// TIA Portal project "000_empty" (V21)

(* hardware
DEVICE "PLC_1"  S7-1500 station
   slot 0: "Rail_0"  Rack  6ES7 590-1***0-0AA0
   slot 1: "PLC_1"  CPU 1513-1 PN  6ES7 513-1AL02-0AB0  V2.9
      slot 3: "CPU display_1"  6ES7591-1AA00-0AA0
      slot 32768: "PROFINET interface_1"  X1
         slot 32769: "Port_1"  X1 P1
         slot 32770: "Port_2"  X1 P2
      slot 34817: "Virtual CP interface port_1"  Virtual CP interface port  Virtual CP interface port
*)

// ===== PLC "PLC_1"  CPU 1513-1 PN =====

VAR_GLOBAL   // PLC tag table "Default tag table"
   "tBool" AT %M0.0 : Bool;
   "tBool2" AT %M0.1 : Bool;
   "tInt" AT %MW2 : Int;
   "tDInt" AT %MD4 : DInt;
   "tReal" AT %MD8 : Real;
   "tWord" AT %MW12 : Word;
   "tByte" AT %MB14 : Byte;
   "tDWord" AT %MD16 : DWord;
   "tTime" AT %MD20 : Time;
   "tIn" AT %I0.0 : Bool;
   "tOut" AT %Q0.0 : Bool;
   "tUInt" AT %MW24 : UInt;
   "tLReal" AT %MD26 : LReal;
   "Tag_1" AT %MW100 : Word;
   "Tag_2" AT %M10.3 : Bool;
   "Tag_3" AT %Q1.0 : Bool;
   "Tag_4" AT %I1.0 : Bool;
   "Tag_5" AT %MD104 : DWord;
   "Tag_6" AT %MB110 : Byte;
   "Tag_7" AT %IW0 : Word;
   "Tag_8" AT %QW0 : Word;
END_VAR

VAR_GLOBAL CONSTANT   // PLC tag table "Default tag table"
   "MAX_COUNT" : Int := 100;
   "GAIN" : Real := 2.5;
   "TXT" : String := 'abc';
END_VAR

TYPE "UDT_Motor"
   STRUCT
      Running : Bool;   // Motor on
      Speed : Real := 1500.0;   // Speed setpoint
      Count : Int := 7;
   END_STRUCT;
END_TYPE

DATA_BLOCK "DB_Global"   // DB1
{ S7_Optimized_Access := 'TRUE' }
   VAR
      xBool : Bool := TRUE;   // Bool comment
      iInt : Int := 42;
      rReal : Real := 3.5;   // Real comment
      aInt : Array[0..3] of Int;
      sData : Struct
         "a" : Bool;
         "b" : DInt := -5;
      END_STRUCT;
   END_VAR
BEGIN
   aInt[1] := 11;
END_DATA_BLOCK

DATA_BLOCK "FB_Empty_DB"   // DB2
{ S7_Optimized_Access := 'TRUE' }
VERSION : 0.1
// stored: InstanceOfName FB_Empty
"FB_Empty"
BEGIN
END_DATA_BLOCK

DATA_BLOCK "DB_Motor"   // DB4
{ S7_Optimized_Access := 'TRUE' }
   VAR
      motor : "UDT_Motor";
   END_VAR
BEGIN
   motor.Speed := 750.0;
END_DATA_BLOCK

DATA_BLOCK "FB_Iface_DB"   // DB5
{ S7_Optimized_Access := 'TRUE' }
VERSION : 0.1
// stored: InstanceOfName FB_Iface
"FB_Iface"
BEGIN
   stInt := 99;
   stBool := TRUE;
END_DATA_BLOCK

DATA_BLOCK "DB_Std"   // DB6
{ S7_Optimized_Access := 'FALSE' }
   VAR
      x : Bool;
      i : Int;
      d : DInt;
      r : Real;
      "by" : Byte;
   END_VAR
BEGIN
END_DATA_BLOCK

DATA_BLOCK "DB_Arr"   // DB7
{ S7_Optimized_Access := 'FALSE' }
   VAR
      "a" : Array[0..9] of Int;
      "b" : Array[0..9] of Int;
      w : Array[0..3] of Word;
      r : Array[0..3] of Real;
      "by" : Array[0..7] of Byte;
      bits : Array[0..15] of Bool;
   END_VAR
BEGIN
END_DATA_BLOCK

// folder: BlockGroup_1

DATA_BLOCK "DB_InGroup"   // DB3
{ S7_Optimized_Access := 'TRUE' }
   VAR
      wWord : Word := 16#00FF;
   END_VAR
BEGIN
END_DATA_BLOCK

// folder: (top level)

FUNCTION_BLOCK "FB_Empty"   // FB1, SCL
{ S7_Optimized_Access := 'TRUE' }
VERSION : 0.1
BEGIN
END_FUNCTION_BLOCK

FUNCTION_BLOCK "FB_Iface"   // FB2, SCL
{ S7_Optimized_Access := 'TRUE' }
VERSION : 0.1
   VAR_INPUT
      iBool : Bool;   // Input bool
      iInt : Int;   // Input int
      iReal : Real;   // Input real
      iArr : Array[0..3] of Int;   // Input array
      iMotor : "UDT_Motor";   // Input UDT
   END_VAR
   VAR_OUTPUT
      oBool : Bool;   // Output bool
      oInt : Int;   // Output int
   END_VAR
   VAR_IN_OUT
      ioReal : Real;   // InOut real
   END_VAR
   VAR
      stInt : Int := 42;   // Static int
      stBool : Bool;   // Static bool comment
   END_VAR
   VAR_TEMP
      tInt : Int;   // Temp int
   END_VAR
   VAR CONSTANT
      cInt : Int := 7;   // Constant int
   END_VAR
BEGIN
   #tInt := #iInt + #cInt;
           #oInt := #tInt;
           #oBool := #iBool;
           #ioReal := #ioReal + #iReal;
END_FUNCTION_BLOCK

FUNCTION_BLOCK "FB_SclCalls"   // FB3, SCL
{ S7_Optimized_Access := 'TRUE' }
VERSION : 0.1
   VAR_INPUT
      start : Bool;
      pt : Time;
   END_VAR
   VAR_OUTPUT
      q : Bool;
      cnt : Int;
   END_VAR
   VAR
      tonInst : TON_TIME;
      tofInst : TOF_TIME;
      tpInst : TP_TIME;
      ctuInst : CTU_INT;
      trig : R_TRIG;
      ftrig : F_TRIG;
      "counter" : Int;
      ifc : "FB_Iface";
   END_VAR
   VAR_TEMP
      r : Real;
      "b" : Bool;
      res : Int;
      tot : Int;
   END_VAR
BEGIN
   #tonInst(IN := #start, PT := #pt);
   #q := #tonInst.Q;
   #tofInst(IN := #start, PT := T#2s);
   #tpInst(IN := #start, PT := #pt, Q => #b);
   #ctuInst(CU := #start, R := FALSE, PV := 10);
   #cnt := #ctuInst.CV;
   #trig(CLK := #start);
   IF #trig.Q THEN
       #counter := 0;
   END_IF;
   #ftrig(CLK := #start);
   #b := #ftrig.Q;
   #ifc(iBool := TRUE, iInt := 2, iReal := 1.0, ioReal := #r);
   #cnt := #ifc.oInt;
   "FB_Iface_DB"(iBool := #start, iInt := #cnt, iReal := #r, ioReal := #r, oInt => #cnt);
   "FC_SclOps"();
   #res := "FC_SclCtl"(n := 5, flag := TRUE, total => #tot);
   #res := "FC_SclCtl"(n := #res, flag := #b, total => #tot);
END_FUNCTION_BLOCK

FUNCTION_BLOCK "FB_SclLocal"   // FB4, SCL
{ S7_Optimized_Access := 'TRUE' }
VERSION : 0.1
   VAR_INPUT
      start : Bool;
   END_VAR
   VAR_IN_OUT
      io : Int;
   END_VAR
   VAR
      "counter" : Int;
      arr : Array[0..9] of Int;
      arr2 : Array[1..3, 1..4] of Real;
      mot : "UDT_Motor";
      st : Struct
         "a" : Int;
         "b" : Real;
         c : Array[0..2] of Bool;
      END_STRUCT;
   END_VAR
   VAR_TEMP
      i : Int;
   END_VAR
BEGIN
   #arr[0] := 1;
   #arr[#i] := #arr[#i + 1] + #io;
   #arr2[2, 3] := 1.5;
   #st.a := 10;
   #st.b := #st.a;
   #st.c[1] := TRUE;
   #mot.Speed := 100.0;
   #mot.Running := #st.c[0];
   #counter += 1;
   #io := #counter;
END_FUNCTION_BLOCK

FUNCTION_BLOCK "FB_Lad_ex005"   // FB5, LAD
{ S7_Optimized_Access := 'TRUE' }
VERSION : 0.1
   VAR_INPUT
      v_in1 : DTL;
      v_in2 : DTL;
      v_out : Time;
   END_VAR
BEGIN

REGION Network 1: T_DIFF - Time difference
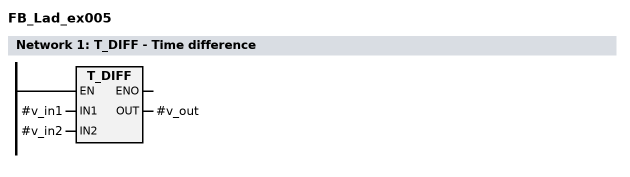
   #v_out := T_DIFF(IN1 := #v_in1, IN2 := #v_in2);
END_REGION
END_FUNCTION_BLOCK

FUNCTION_BLOCK "FB_Lad_ex007"   // FB6, LAD
{ S7_Optimized_Access := 'TRUE' }
VERSION : 0.1
   VAR_INPUT
      v_in : DTL;
      v_ret_val : Int;
   END_VAR
BEGIN

REGION Network 1: WR_SYS_T - Set time-of-day
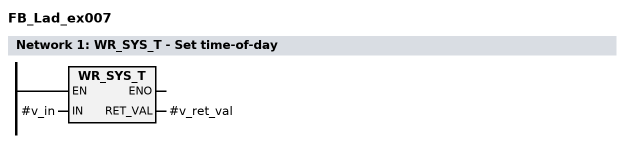
   #v_ret_val := WR_SYS_T(IN := #v_in);
END_REGION
END_FUNCTION_BLOCK

FUNCTION_BLOCK "FB_Lad_ex008"   // FB7, LAD
{ S7_Optimized_Access := 'TRUE' }
VERSION : 0.1
   VAR_INPUT
      v_ret_val : Int;
   END_VAR
   VAR_OUTPUT
      v_out : DTL;
   END_VAR
BEGIN

REGION Network 1: RD_SYS_T - Read time-of-day
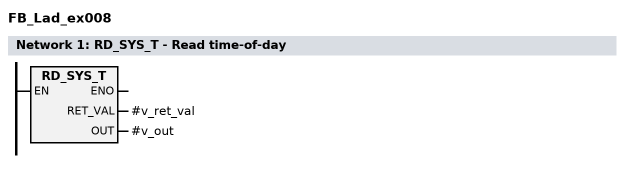
   #v_ret_val := RD_SYS_T(OUT => #v_out);
END_REGION
END_FUNCTION_BLOCK

FUNCTION_BLOCK "FB_Lad_ex009"   // FB8, LAD
{ S7_Optimized_Access := 'TRUE' }
VERSION : 0.1
   VAR_INPUT
      v_ret_val : Int;
   END_VAR
   VAR_OUTPUT
      v_out : DTL;
   END_VAR
BEGIN

REGION Network 1: RD_LOC_T - Read local time
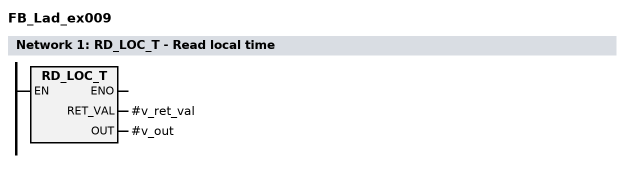
   #v_ret_val := RD_LOC_T(OUT => #v_out);
END_REGION
END_FUNCTION_BLOCK

FUNCTION_BLOCK "FB_Lad_ex012"   // FB9, LAD
{ S7_Optimized_Access := 'TRUE' }
VERSION : 0.1
   VAR_OUTPUT
      v_ret_val : Int;
   END_VAR
BEGIN

REGION Network 1: SNC_RTCB - Synchronize slave clocks
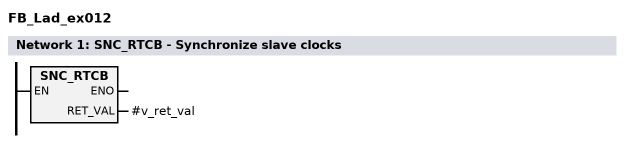
   #v_ret_val := SNC_RTCB();
END_REGION
END_FUNCTION_BLOCK

FUNCTION_BLOCK "FB_Lad_ex013"   // FB10, LAD
{ S7_Optimized_Access := 'TRUE' }
VERSION : 0.1
   VAR_INPUT
      v_ret_val : Time;
   END_VAR
BEGIN

REGION Network 1: TIME_TCK - Read time counter
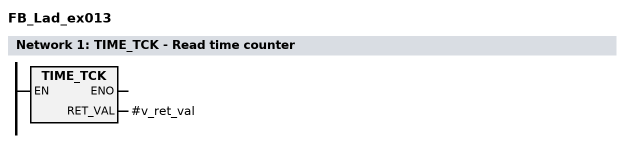
   #v_ret_val := TIME_TCK();
END_REGION
END_FUNCTION_BLOCK

FUNCTION_BLOCK "FB_Lad_ex014"   // FB11, LAD
{ S7_Optimized_Access := 'TRUE' }
VERSION : 0.1
   VAR_INPUT
      v_nr : Rtm;
      v_mode : Byte;
      v_pv : DInt;
      v_ret_val : Int;
   END_VAR
   VAR_OUTPUT
      v_cq : Bool;
      v_cv : DInt;
   END_VAR
BEGIN

REGION Network 1: RTM - Runtime meters
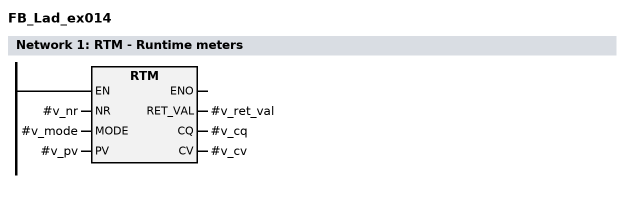
   #v_ret_val := RTM(NR := #v_nr, MODE := #v_mode, PV := #v_pv, CQ => #v_cq, CV => #v_cv);
END_REGION
END_FUNCTION_BLOCK

FUNCTION_BLOCK "FB_Lad_ex015"   // FB12, LAD
{ S7_Optimized_Access := 'TRUE' }
VERSION : 0.1
   VAR_INPUT
      v_in : String;
   END_VAR
   VAR_OUTPUT
      v_out : String;
   END_VAR
BEGIN

REGION Network 1: S_MOVE - Move character string
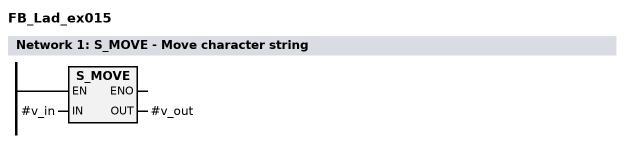
   RUNG wire#powerrail
      S_Move(in := #v_in, out => #v_out)
   END_RUNG
   // the same network as SCL:
   #v_out := #v_in;
END_REGION
END_FUNCTION_BLOCK

FUNCTION_BLOCK "FB_Lad_ex038"   // FB13, LAD
{ S7_Optimized_Access := 'TRUE' }
   VAR_INPUT
      v_size : DInt;
   END_VAR
   VAR_OUTPUT
      v_out : WString;
   END_VAR
BEGIN

REGION Network 1: GetInstanceName - Read out name of the read instance
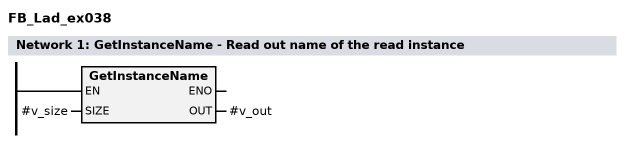
   // no SCL statement known for GetInstanceName: written as a call
   #v_out := GetInstanceName(size := #v_size);
END_REGION
END_FUNCTION_BLOCK

FUNCTION_BLOCK "FB_Lad_ex039"   // FB14, LAD
{ S7_Optimized_Access := 'TRUE' }
   VAR_INPUT
      v_size : DInt;
   END_VAR
   VAR_OUTPUT
      v_out : WString;
   END_VAR
BEGIN

REGION Network 1: GetInstancePath - Query composite global name of the block instance
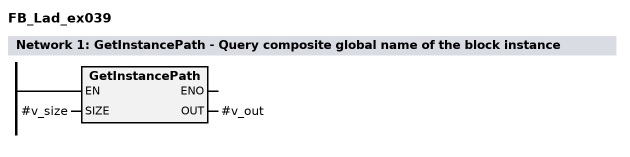
   // no SCL statement known for GetInstancePath: written as a call
   #v_out := GetInstancePath(size := #v_size);
END_REGION
END_FUNCTION_BLOCK

FUNCTION_BLOCK "FB_Lad_ex040"   // FB15, LAD
{ S7_Optimized_Access := 'TRUE' }
   VAR_INPUT
      v_size : DInt;
   END_VAR
   VAR_OUTPUT
      v_ret_val : WString;
   END_VAR
BEGIN

REGION Network 1: GetBlockName - Read out name of the block
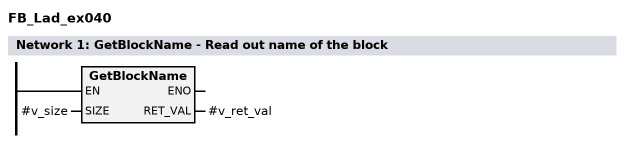
   // no SCL statement known for GetBlockName: written as a call
   #v_ret_val := GetBlockName(size := #v_size);
END_REGION
END_FUNCTION_BLOCK

FUNCTION_BLOCK "FB_Lad_ex041"   // FB16, LAD
{ S7_Optimized_Access := 'TRUE' }
   VAR_INPUT
      v_part : Pip;
      v_ret_val : Int;
   END_VAR
   VAR_OUTPUT
      v_fladdr : Word;
   END_VAR
BEGIN

REGION Network 1: UPDAT_PI - Update the process image inputs
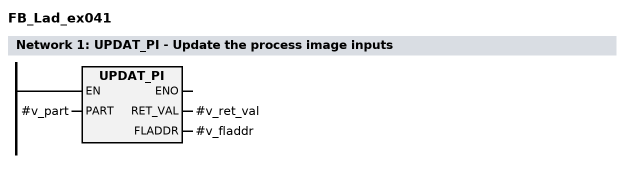
   #v_ret_val := UPDAT_PI(PART := #v_part, FLADDR => #v_fladdr);
END_REGION
END_FUNCTION_BLOCK

FUNCTION_BLOCK "FB_Lad_ex042"   // FB17, LAD
{ S7_Optimized_Access := 'TRUE' }
   VAR_INPUT
      v_part : Pip;
      v_ret_val : Int;
   END_VAR
   VAR_OUTPUT
      v_fladdr : Word;
   END_VAR
BEGIN

REGION Network 1: UPDAT_PO - Update the process image outputs
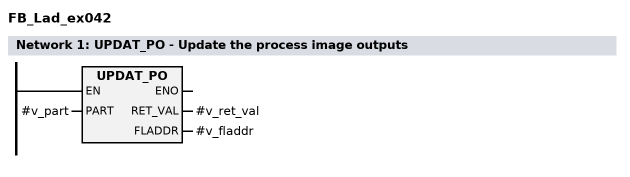
   #v_ret_val := UPDAT_PO(PART := #v_part, FLADDR => #v_fladdr);
END_REGION
END_FUNCTION_BLOCK

FUNCTION_BLOCK "FB_Lad_ex043"   // FB18, LAD
{ S7_Optimized_Access := 'TRUE' }
   VAR_INPUT
      v_part : Pip;
      v_ret_val : Int;
   END_VAR
   VAR_OUTPUT
      v_fladdr : Word;
   END_VAR
BEGIN

REGION Network 1: SYNC_PI - Synchronize the process image inputs
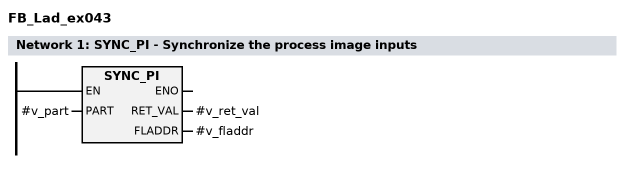
   #v_ret_val := SYNC_PI(PART := #v_part, FLADDR => #v_fladdr);
END_REGION
END_FUNCTION_BLOCK

FUNCTION_BLOCK "FB_Lad_ex044"   // FB19, LAD
{ S7_Optimized_Access := 'TRUE' }
   VAR_INPUT
      v_part : Pip;
      v_ret_val : Int;
   END_VAR
   VAR_OUTPUT
      v_fladdr : Word;
   END_VAR
BEGIN

REGION Network 1: SYNC_PO - Synchronize the process image outputs
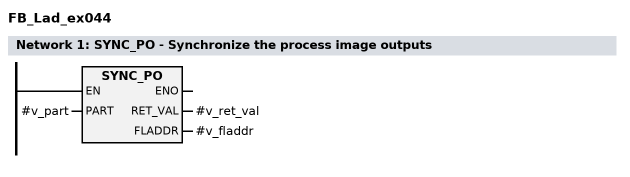
   #v_ret_val := SYNC_PO(PART := #v_part, FLADDR => #v_fladdr);
END_REGION
END_FUNCTION_BLOCK

FUNCTION_BLOCK "FB_Lad_ex056"   // FB20, LAD
{ S7_Optimized_Access := 'TRUE' }
   VAR_INPUT
      v_req : Bool;
      v_mode : USInt;
      v_laddr : Hw_Device;
      v_ret_val : Int;
   END_VAR
   VAR_OUTPUT
      v_busy : Bool;
   END_VAR
BEGIN

REGION Network 1: D_ACT_DP - Activate/deactivate DP slaves
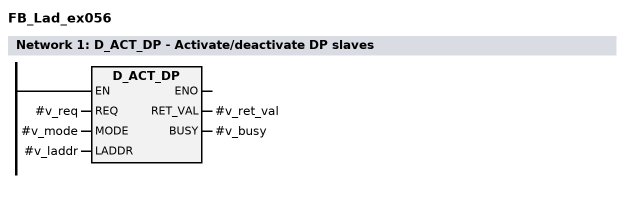
   #v_ret_val := D_ACT_DP(REQ := #v_req, MODE := #v_mode, LADDR := #v_laddr, BUSY => #v_busy);
END_REGION
END_FUNCTION_BLOCK

FUNCTION_BLOCK "FB_Lad_ex061"   // FB21, LAD
{ S7_Optimized_Access := 'TRUE' }
   VAR_INPUT
      v_laddr : Hw_Io;
      v_record : Variant;
      v_ret_val : Int;
   END_VAR
BEGIN

REGION Network 1: DPWR_DAT - Write consistent data of a DP standard slave
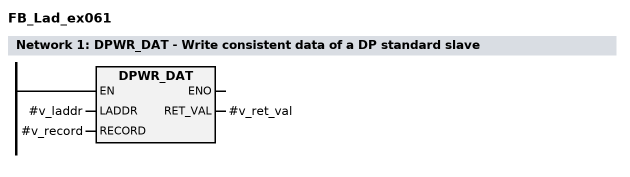
   #v_ret_val := DPWR_DAT(LADDR := #v_laddr, RECORD := #v_record);
END_REGION
END_FUNCTION_BLOCK

FUNCTION_BLOCK "FB_Lad_ex064"   // FB22, LAD
{ S7_Optimized_Access := 'TRUE' }
   VAR_INPUT
      v_req : Bool;
      v_laddr : Hw_Interface;
      v_group : Byte;
      v_mode : Byte;
      v_ret_val : Int;
   END_VAR
   VAR_OUTPUT
      v_busy : Bool;
   END_VAR
BEGIN

REGION Network 1: DPSYC_FR - Synchronize DP slaves / Freeze inputs
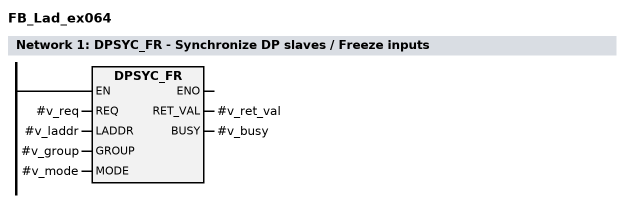
   #v_ret_val := DPSYC_FR(REQ := #v_req, LADDR := #v_laddr, GROUP := #v_group, MODE := #v_mode, BUSY => #v_busy);
END_REGION
END_FUNCTION_BLOCK

FUNCTION_BLOCK "FB_Lad_ex066"   // FB23, LAD
{ S7_Optimized_Access := 'TRUE' }
   VAR_INPUT
      v_req : Bool;
      v_r : Bool;
      v_dp_id : Hw_IoSystem;
      v_ret_val : Int;
   END_VAR
   VAR_OUTPUT
      v_busy : Bool;
      v_dpr : Byte;
      v_dpri : Byte;
   END_VAR
BEGIN

REGION Network 1: DP_TOPOL - Determine topology for DP master system
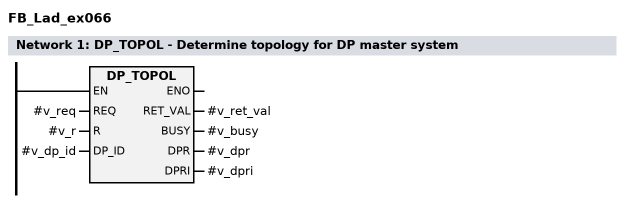
   #v_ret_val := DP_TOPOL(REQ := #v_req,
                          R := #v_r,
                          DP_ID := #v_dp_id,
                          BUSY => #v_busy,
                          DPR => #v_dpr,
                          DPRI => #v_dpri);
END_REGION
END_FUNCTION_BLOCK

FUNCTION_BLOCK "FB_Lad_ex099"   // FB24, LAD
{ S7_Optimized_Access := 'TRUE' }
   VAR_INPUT
      v_req : Bool;
      v_laddr : Hw_Io;
      v_recnum : Byte;
      v_ret_val : Int;
   END_VAR
   VAR_OUTPUT
      v_busy : Bool;
   END_VAR
BEGIN

REGION Network 1: WR_DPARM - Transfer data record
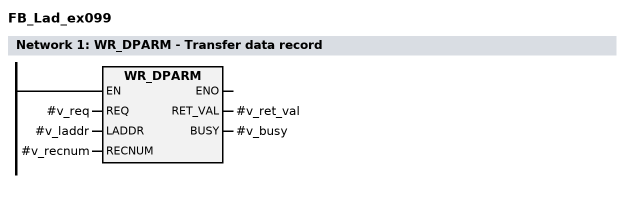
   #v_ret_val := WR_DPARM(REQ := #v_req, LADDR := #v_laddr, RECNUM := #v_recnum, BUSY => #v_busy);
END_REGION
END_FUNCTION_BLOCK

FUNCTION_BLOCK "FB_Lad_ex100"   // FB25, LAD
{ S7_Optimized_Access := 'TRUE' }
   VAR_INPUT
      v_ob_nr : OB_Att;
      v_event : Event_Att;
      v_add : Bool;
      v_ret_val : Int;
   END_VAR
BEGIN

REGION Network 1: ATTACH - Attach an OB to an interrupt event
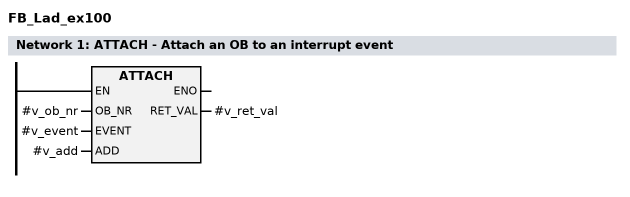
   #v_ret_val := ATTACH(OB_NR := #v_ob_nr, EVENT := #v_event, ADD := #v_add);
END_REGION
END_FUNCTION_BLOCK

FUNCTION_BLOCK "FB_Lad_ex101"   // FB26, LAD
{ S7_Optimized_Access := 'TRUE' }
   VAR_INPUT
      v_ob_nr : OB_Att;
      v_event : Event_Att;
      v_ret_val : Int;
   END_VAR
BEGIN

REGION Network 1: DETACH - Detach an OB from an interrupt event
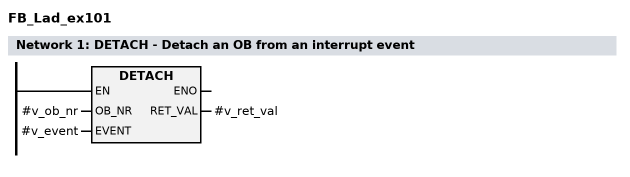
   #v_ret_val := DETACH(OB_NR := #v_ob_nr, EVENT := #v_event);
END_REGION
END_FUNCTION_BLOCK

FUNCTION_BLOCK "FB_Lad_ex102"   // FB27, LAD
{ S7_Optimized_Access := 'TRUE' }
   VAR_INPUT
      v_ob_nr : OB_Cyclic;
      v_cycle : UDInt;
      v_phase : UDInt;
      v_ret_val : Int;
   END_VAR
BEGIN

REGION Network 1: SET_CINT - Set cyclic interrupt parameters
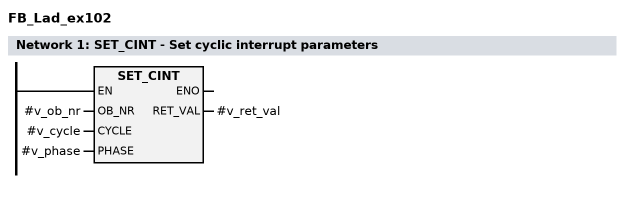
   #v_ret_val := SET_CINT(OB_NR := #v_ob_nr, CYCLE := #v_cycle, PHASE := #v_phase);
END_REGION
END_FUNCTION_BLOCK

FUNCTION_BLOCK "FB_Lad_ex103"   // FB28, LAD
{ S7_Optimized_Access := 'TRUE' }
   VAR_INPUT
      v_ob_nr : Int;
      v_ret_val : Int;
   END_VAR
   VAR_OUTPUT
      v_cycle : UDInt;
      v_phase : UDInt;
      v_status : Word;
   END_VAR
BEGIN

REGION Network 1: QRY_CINT - Query cyclic interrupt parameters
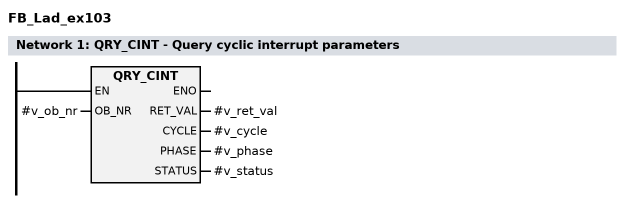
   #v_ret_val := QRY_CINT(OB_NR := #v_ob_nr, CYCLE => #v_cycle, PHASE => #v_phase, STATUS => #v_status);
END_REGION
END_FUNCTION_BLOCK

FUNCTION_BLOCK "FB_Lad_ex104"   // FB29, LAD
{ S7_Optimized_Access := 'TRUE' }
   VAR_INPUT
      v_ob_nr : OB_Tod;
      v_sdt : Date_And_Time;
      v_period : Word;
      v_ret_val : Int;
   END_VAR
BEGIN

REGION Network 1: SET_TINT - Set time-of-day interrupt
